(* IEC 61131-3 sources: Lasal-MCP/examples/SampleSource/5_ClassInputOutputSolution/Stations/MachineControl/MachineControl/Class/PcComponentsRadio, 1 file *)

(* ---- PcComponentsRadio.st ---- *)
(*!
<Class
	Name               = "PcComponentsRadio"
	Revision           = "0.0"
	RealtimeTask       = "false"
	CyclicTask         = "false"
	BackgroundTask     = "false"
	Sigmatek           = "false"
	OSInterface        = "false"
	HighPriority       = "false"
	Automatic          = "false"
	UpdateMode         = "Prescan"
	SharedCommandTable = "true"
	Objectsize         = "(512,120)">
	<Channels>
		<Server Name="MyComponents" Visualized="true" Initialize="false" WriteProtected="false" Retentive="false"/>
		<Client Name="_Radio321" Required="true" Internal="true"/>
	</Channels>
	<Network Name="PcComponentsRadio">
		<!-- List of Components in this network -->
		<Components>
			<Object
				Name       = "_Radio321"
				Class      = "_Radio32"
				Position   = "(150,330)"
				Visualized = "true"
				Remotely   = "true">
				<Channels>
					<Server Name="Data"/>
				</Channels>
			</Object>
		</Components>
		<Comments>
		</Comments>
		<!-- List of Connections in this network -->
		<Connections>
			<Connection Source="this._Radio321" Destination="_Radio321.Data"/>
		</Connections>
		<!-- Headerfiles -->
		<Options>
		</Options>
	</Network>
</Class>
*)
PcComponentsRadio : CLASS
	TYPE
	  t_PC_COMPONENTS : BDINT  //! <Type Public="true" Name="t_PC_COMPONENTS"/>
	  [
	    1 Mouse,
	    2 Keyboard,
	    3 USB,
	    4 Monitor,
	    5 Bit5,
	    6 Bit6,
	    7 Bit7,
	    8 Bit8,
	    9 Bit9,
	    10 Bit10,
	    11 Bit11,
	    12 Bit12,
	    13 Bit13,
	    14 Bit14,
	    15 Bit15,
	    16 Bit16,
	    17 Bit17,
	    18 Bit18,
	    19 Bit19,
	    20 Bit20,
	    21 Bit21,
	    22 Bit22,
	    23 Bit23,
	    24 Bit24,
	    25 Bit25,
	    26 Bit26,
	    27 Bit27,
	    28 Bit28,
	    29 Bit29,
	    30 Bit30,
	    31 Bit31,
	    32 Bit32,
	  ];
	END_TYPE
  //Servers:
	MyComponents 	: SvrChCmd_t_PC_COMPONENTS_PTofCls_PcComponentsRadio;
  //Clients:
	_Radio321 	: CltChCmd__Radio32;
  //Variables:
  //Functions:

	FUNCTION VIRTUAL GLOBAL MyComponents::Write
		VAR_INPUT
			input (EAX) 	: PcComponentsRadio::t_PC_COMPONENTS;
		END_VAR
		VAR_OUTPUT
			result (EAX) 	: PcComponentsRadio::t_PC_COMPONENTS;
		END_VAR;
  //Tables:
	FUNCTION @STD
		VAR_OUTPUT
			ret_code	: CONFSTATES;
		END_VAR;
	FUNCTION GLOBAL TAB @CT_;
END_CLASS;

#pragma using _Radio32

FUNCTION VIRTUAL GLOBAL PcComponentsRadio::MyComponents::Write
	VAR_INPUT
		input (EAX) 	: PcComponentsRadio::t_PC_COMPONENTS;
	END_VAR
	VAR_OUTPUT
		result (EAX) 	: PcComponentsRadio::t_PC_COMPONENTS;
	END_VAR

	MyComponents := _Radio321.Data.Write(input:=input);

	result := MyComponents;

END_FUNCTION
